(* IEC 61131-3 sources: XPGAnalyser/projets/ihm/project/ihm/fonctions, 1 file *)

(* ---- 0031-Fonction.st ---- *)
(* Fonction *)
VAR_INPUT
    Entree : REAL;
END_VAR
VAR_TEMP
    Resultat : REAL;
END_VAR

Resultat := Entree;
Fonction := Resultat;
